Fanuc KAREL source: KB00122.KL

PROGRAM KB00122
%NOLOCKGROUP
%ENVIRONMENT FDEV
VAR
  P1: STRING[80]
  P2: INTEGER
BEGIN
  P1 = 'A'
  P2 = 1
  MOUNT_DEV(P1, P2)
END KB00122
